TYPE ST_ConveyorConfig :
STRUCT
    enabled : BOOL := TRUE;
    speed : LREAL := 0.75;
END_STRUCT
END_TYPE

(* stored: Version 1.1.0.1, ProductVersion 3.1 *)
